(* IEC 61131-3 sources: llm-plc-st-eval/data/processed_definitivo/gemini-3.1-pro-preview/I7/zero_shot, 3 files *)

(* ---- ejec_1.st ---- *)
FUNCTION_BLOCK FB_Duplex
VAR_INPUT
    demanda : BOOL; (* Señal de petición de funcionamiento *)
    falla1  : BOOL; (* Señal de falla de la bomba 1 *)
    falla2  : BOOL; (* Señal de falla de la bomba 2 *)
END_VAR
VAR_OUTPUT
    bomba1   : BOOL; (* Comando de marcha para la bomba 1 *)
    bomba2   : BOOL; (* Comando de marcha para la bomba 2 *)
    almFalla : BOOL; (* Alarma activa si la bomba principal falla durante la demanda *)
END_VAR
VAR
    demandaAnt     : BOOL := FALSE; (* Memoria del estado anterior de la demanda *)
    turnoBomba1    : BOOL := TRUE;  (* TRUE = Bomba 1 principal, FALSE = Bomba 2 principal *)
    primerArranque : BOOL := TRUE;  (* Bandera para forzar bomba 1 en la primera demanda *)
END_VAR

(* Detección de flanco de subida en la demanda para alternar el turno *)
IF demanda AND NOT demandaAnt THEN
    IF primerArranque THEN
        turnoBomba1 := TRUE;
        primerArranque := FALSE;
    ELSE
        turnoBomba1 := NOT turnoBomba1;
    END_IF;
END_IF;
demandaAnt := demanda;

(* Inicialización de salidas (estado de reposo) *)
bomba1   := FALSE;
bomba2   := FALSE;
almFalla := FALSE;

(* Lógica de operación cuando hay demanda activa *)
IF demanda THEN
    IF turnoBomba1 THEN
        (* Turno: Bomba 1 es la principal *)
        IF NOT falla1 THEN
            bomba1 := TRUE;
        ELSE
            almFalla := TRUE; (* Falla la principal, se activa alarma *)
            IF NOT falla2 THEN
                bomba2 := TRUE; (* Entra la bomba 2 de respaldo *)
            END_IF;
        END_IF;
    ELSE
        (* Turno: Bomba 2 es la principal *)
        IF NOT falla2 THEN
            bomba2 := TRUE;
        ELSE
            almFalla := TRUE; (* Falla la principal, se activa alarma *)
            IF NOT falla1 THEN
                bomba1 := TRUE; (* Entra la bomba 1 de respaldo *)
            END_IF;
        END_IF;
    END_IF;
END_IF;

END_FUNCTION_BLOCK

(* ---- ejec_2.st ---- *)
FUNCTION_BLOCK FB_Duplex
VAR_INPUT
    demanda : BOOL; (* Señal de demanda del sistema *)
    falla1  : BOOL; (* Señal de falla de la bomba 1 *)
    falla2  : BOOL; (* Señal de falla de la bomba 2 *)
END_VAR
VAR_OUTPUT
    bomba1   : BOOL; (* Comando de marcha para la bomba 1 *)
    bomba2   : BOOL; (* Comando de marcha para la bomba 2 *)
    almFalla : BOOL; (* Alarma de falla de la bomba principal *)
END_VAR
VAR
    flancoDemanda   : R_TRIG; (* Detector de flanco de subida *)
    bomba1Principal : BOOL := FALSE; (* Inicia en FALSE para cambiar a TRUE en la 1ra demanda *)
END_VAR

(* Detectar transición de FALSE a TRUE en la demanda *)
flancoDemanda(CLK := demanda);

(* Alternar el rol de bomba principal en cada nueva demanda *)
IF flancoDemanda.Q THEN
    bomba1Principal := NOT bomba1Principal;
END_IF;

(* Lógica de control de bombas y alarma *)
IF demanda THEN
    IF bomba1Principal THEN
        (* Ciclo donde Bomba 1 es la principal *)
        bomba1   := NOT falla1;
        bomba2   := falla1 AND NOT falla2; (* Respaldo si la principal falla y respaldo está OK *)
        almFalla := falla1;                (* Alarma activa solo por falla de la principal *)
    ELSE
        (* Ciclo donde Bomba 2 es la principal *)
        bomba2   := NOT falla2;
        bomba1   := falla2 AND NOT falla1; (* Respaldo si la principal falla y respaldo está OK *)
        almFalla := falla2;                (* Alarma activa solo por falla de la principal *)
    END_IF;
ELSE
    (* Si no hay demanda, se detienen las bombas y se apaga la alarma *)
    bomba1   := FALSE;
    bomba2   := FALSE;
    almFalla := FALSE;
END_IF;
END_FUNCTION_BLOCK

(* ---- ejec_3.st ---- *)
FUNCTION_BLOCK FB_Duplex
VAR_INPUT
    demanda : BOOL; // Señal de demanda para arrancar el sistema
    falla1  : BOOL; // Señal de falla activa de la bomba 1
    falla2  : BOOL; // Señal de falla activa de la bomba 2
END_VAR

VAR_OUTPUT
    bomba1   : BOOL; // Comando de operación para la bomba 1
    bomba2   : BOOL; // Comando de operación para la bomba 2
    almFalla : BOOL; // Alarma de falla de la bomba principal con demanda presente
END_VAR

VAR
    rTrigDemanda    : R_TRIG; // Detector de flanco de subida de la demanda
    bomba1Principal : BOOL := TRUE; // Indica si la bomba 1 tiene el rol principal
    primerArranque  : BOOL := TRUE; // Bandera para identificar la primera demanda
END_VAR

// Detección del flanco de subida de la señal de demanda
rTrigDemanda(CLK := demanda);

// Lógica de alternancia en cada nueva demanda
IF rTrigDemanda.Q THEN
    IF primerArranque THEN
        // En la primera demanda tras el arranque, la principal es la bomba 1
        primerArranque := FALSE;
    ELSE
        // En las demandas posteriores, se alterna el rol principal
        bomba1Principal := NOT bomba1Principal;
    END_IF;
END_IF;

// Lógica de control de operación y respaldo
IF demanda THEN
    IF bomba1Principal THEN
        // Bomba 1 es la principal, Bomba 2 es el respaldo
        bomba1   := NOT falla1;
        bomba2   := falla1 AND NOT falla2;
        almFalla := falla1;
    ELSE
        // Bomba 2 es la principal, Bomba 1 es el respaldo
        bomba2   := NOT falla2;
        bomba1   := falla2 AND NOT falla1;
        almFalla := falla2;
    END_IF;
ELSE
    // Al desactivarse la demanda, ambas bombas se detienen y se apaga la alarma
    bomba1   := FALSE;
    bomba2   := FALSE;
    almFalla := FALSE;
END_IF;

END_FUNCTION_BLOCK
